TYPE ST_ConfigXtsLoop :
STRUCT
	(* vo_Config of _FB_ConfigXtsLoop: the gateway writes stStaging and stStaged, reads stStatus and stActive. *)
	stStaging : ST_ConfigStaging;
	stStaged : ST_ConfigXtsLoopParam;
	stStatus : ST_ConfigStatus;
	stActive : ST_ConfigXtsLoopParam; // effective values: the active set while one is valid, else the program values
END_STRUCT
END_TYPE

(* stored: Version 1.1.0.1
   DUT ST_ConfigXtsLoop: Id {eb5169c6-4b3f-4ab4-8c69-147e8b10381a} *)
